Fanuc KAREL source: kf00099.KL

-- PROVISIONAL review KL for V940-1; original PC SHA256 1a2cfe69f2d3e903d336d41b9b29e6341c6ca510a3f114533b46345d17e74e56
-- Incomplete behavior may be omitted. Consult companion uncertainty JSON. Do not deploy.
PROGRAM KF00099
%NOLOCKGROUP
BEGIN
  -- V9_ZERO_TABLE_METADATA_HINT layout=0002_ascii; no indexed target words; source/name/runtime held
  -- UNRESOLVED_PC offsets 5-16; opcodes 2E,23
  -- UNRESOLVED_PC offsets 21-32; opcodes 2E,23
  -- UNRESOLVED_PC offsets 37-63; opcodes 27,27,9D,22,27,9D,31,7E,4A
  -- UNRESOLVED_PC offsets 68-72; opcodes 7F
END KF00099
